(* IEC 61131-3 sources: llm-plc-st-eval/data/definitivo/gemini-3.1-pro-preview/B7/few_shot, 3 files *)

(* ---- ejec_1.st ---- *)
FUNCTION SelBomba : BOOL
VAR_INPUT
    modoAuto : BOOL; (* Modo automatico activo *)
    btnManual : BOOL; (* Boton de mando manual *)
    nivelBajo : BOOL; (* Sensor de nivel bajo *)
END_VAR

(* Seleccion de mando: nivel en automatico, boton en manual *)
SelBomba := (modoAuto AND nivelBajo) OR (NOT modoAuto AND btnManual);
END_FUNCTION

(* ---- ejec_2.st ---- *)
FUNCTION SelBomba : BOOL
VAR_INPUT
    modoAuto : BOOL; (* Modo automatico activo *)
    btnManual : BOOL; (* Boton de mando manual *)
    nivelBajo : BOOL; (* Sensor de nivel bajo *)
END_VAR

(* Logica sin memoria: obedece al sensor en auto o al boton en manual *)
SelBomba := (modoAuto AND nivelBajo) OR (NOT modoAuto AND btnManual);
END_FUNCTION

(* ---- ejec_3.st ---- *)
FUNCTION SelBomba : BOOL
VAR_INPUT
    modoAuto : BOOL; (* Activa el modo automatico *)
    btnManual : BOOL; (* Boton de mando en modo manual *)
    nivelBajo : BOOL; (* Condicion de encendido en modo automatico *)
END_VAR

(* Estado de la bomba segun el modo seleccionado sin memoria *)
SelBomba := (modoAuto AND nivelBajo) OR (NOT modoAuto AND btnManual);
END_FUNCTION
